// TIA Portal V17 export
DATA_BLOCK "MCP_RC_DB2"   // DB9802
{ S7_Optimized_Access := 'TRUE' }
   VAR
      Count : Int := 16#0A;
      Motor : "MCP_RC_UDT";
      Val : Real := 1.50;
   END_VAR
BEGIN
END_DATA_BLOCK
